TYPE E_LightTargetType :
(
    Light,
    Group
);
END_TYPE

(* stored: Version 1.1.0.1, ProductVersion 3.1.4026.20
   DUT E_LightTargetType: Id {D1A10003-0A11-4A11-8A11-000000000003} *)
